Fanuc KAREL source: KA00167.KL

PROGRAM KA00167
%NOLOCKGROUP
VAR
  SRC: ARRAY[4] OF BOOLEAN
  DST: ARRAY[4] OF BYTE
BEGIN
  DST = SRC
END KA00167
